FUNCTION RemovePlusSign : STRING(254)
VAR_INPUT
    inString : STRING(254);
END_VAR

// Preserve the reference behavior: remove only one leading plus sign.
RemovePlusSign := inString;
IF LEFT(inString, 1) = '+' THEN
    RemovePlusSign := RIGHT(inString, LEN(inString) - 1);
END_IF;

END_FUNCTION

(* stored: Version 1.1.0.1
   POU RemovePlusSign: Id {6b09d02e-7105-48ef-aa27-979431561c53}, SpecialFunc None *)
